(* IEC 61131-3 sources: plcassist-cli/packages/volt-lsp-iec/test-corpus/lenze-mid/Device/Plc Logic/Application/Library Manager/L_OEEA_Library, 3.26.4.21 (Lenze), 23 files *)

(* ---- GVL_AXISSIM.gvl ---- *)
VAR_GLOBAL
	FEEDERAXIS : AXIS_REF_SIM := STRUCT(eTraversingRange := 1, lrCycleLength := 1000.0, lrFeedConstant := 1000.0, dwGearNumerator := 100, dwGearDenominator := 1, eMctrlMode := 0, wNoOfHTLPeriods := 128);
END_VAR

(* ---- GVL_VALIDATIONTEST.gvl ---- *)
VAR_GLOBAL
	SCEXECUTETIMEARRAY : scExecuteTimeArray;
	SCMACHINEDATA_BASE : scMachineData_base;
	SCPERFORMANCE_BASE : scPerformance_base;
	ULISTART : ULINT;
	ULIEND : ULINT;
	XPRODUCTIONACTIVE : BOOL := TRUE;
	FBMACHINEPERFORMANCE_BASE : L_OEEA_MachinePerformance_Base;
	FBDOWNTIME_BASE : L_OEEA_Downtime_base;
	FBSHIFTOEEHISTORYALL : L_OEEA_ShiftOEEHistory;
	FBSHIFTOEEHISTORY_BASE : L_OEEA_ShiftOEEHistory_Base;
	FBSHIFTDOWNTIMEHISTORY_BASE : L_OEEA_ShiftDowntimeHistory_base;
	SCPDINTERNAL_BASE : scInternalVar;
	SCPDSHIFTDAYINDEX : scPDShiftData;
	SCPDINTERNALDOWNTIME_BASE : scInternalDownVar;
	SCDOWNTIME_BASE : scDowntime_base;
	SCSHIFTDOWNTIMEHISTORY_BASE : ARRAY [1..3] OF scDowntime_base;
	SCSHIFTHISTORYALL : ARRAY [1..3] OF scPerformance;
	SCPDSHIFTHISTORY_BASE : scVisuShiftHistory_base;
	SCPDPRODUCTIONDATA : scInternalProductionData;
	SCSHIFTVALUES : scCurrentShiftValues;
END_VAR

(* ---- LINE_OEE_GVL_VAR.gvl ---- *)
VAR_GLOBAL
	UINOOFMACHINES : UINT := 60;
	UINOOFHISTORICALWEEKS : UINT := 4;
END_VAR

(* ---- VERSIONCONSTANTS.gvl ---- *)
VAR_GLOBAL
	GC_BYAMOUNTOFGENERALDATA : BYTE := 50;
	GC_BYAMOUNTDOWNTIMEERRORS : BYTE := 10;
	GC_IFILTERSAMPLES : INT := 20;
END_VAR

(* ---- CALENDAR_WEEK.fun ---- *)
FUNCTION CALENDAR_WEEK : UINT
VAR_INPUT
	DTEXTDT : DATE_AND_TIME;
END_VAR
END_FUNCTION

(* ---- EXECUTIONTIME.fun ---- *)
FUNCTION EXECUTIONTIME : BOOL
VAR_INPUT
	SFBSTR : STRING;
	ULISTART : ULINT;
	ULIEND : ULINT;
END_VAR
VAR_IN_OUT
	AEXECUTION : scExecuteTime;
END_VAR
END_FUNCTION

(* ---- L_OEEA_CUSTOMIZABLE_COPYSTRUCT.fun ---- *)
FUNCTION L_OEEA_CUSTOMIZABLE_COPYSTRUCT : BOOL
VAR_INPUT
	PBYSOURCE : POINTER TO BYTE;
	PBYTARGET : POINTER TO BYTE;
	UISIZESOURCE : UINT;
	UISIZETARGET : UINT;
END_VAR
END_FUNCTION

(* ---- LRAXISPOSCOUNT.fun ---- *)
FUNCTION LRAXISPOSCOUNT : LREAL
VAR_INPUT
	LRAXISPOS : LREAL;
END_VAR
VAR_IN_OUT
	SCAXISPOSCOUNT : scAxisPosCount;
END_VAR
END_FUNCTION

(* ---- GLOBALTEXTLIST.fb ---- *)
FUNCTION_BLOCK GLOBALTEXTLIST
VAR
	M_TEXTLISTFILE : STRING(255);
	_STNAMESPACE : STRING;
END_VAR
END_FUNCTION_BLOCK

(* ---- IMAGEPOOL_AXIS_REF_SIM.fb ---- *)
FUNCTION_BLOCK IMAGEPOOL_AXIS_REF_SIM
VAR
	M_STNAMESPACE : STRING(80);
	M_STHELPVARID : STRING;
	M_STHELPVARPATH : STRING(255);
	M_STHELP : STRING;
	M_REGISTERIMAGES : BOOL := TRUE;
END_VAR
END_FUNCTION_BLOCK

METHOD FB_INIT : BOOL
VAR_INPUT
	BINITRETAINS : BOOL;
	BINCOPYCODE : BOOL;
END_VAR
END_METHOD

METHOD FB_REINIT : BOOL
END_METHOD

METHOD FB_EXIT : BOOL
VAR_INPUT
	BINCOPYCODE : BOOL;
END_VAR
END_METHOD

(* ---- L_MC1A_BASICACTUATINGSPEED.fb ---- *)
FUNCTION_BLOCK L_MC1A_BASICACTUATINGSPEED
VAR_INPUT
	XREGULATORON : BOOL;
	XRESETERROR : BOOL;
	XSETDRIVEQSP : BOOL;
	XENABLESETVEL : BOOL;
	XINVERTDIRECTION : BOOL;
	LRSETVEL : LREAL := 300.0;
	LRSETACC : LREAL := 100.0;
	LRSETDEC : LREAL := 100.0;
END_VAR
VAR_OUTPUT
	XERROR : BOOL;
	XBUSY : BOOL;
	EERRORID : L_IE1A_ErrorID;
	XCOMMUNICATIONOK : BOOL;
	XAXISREADY : BOOL;
	XAXISENABLED : BOOL;
	XDRIVEWARNING : BOOL;
	XDRIVEERROR : BOOL;
	DWDRIVEERRORID : DWORD;
	XDRIVEQSPACTIVE : BOOL;
	LRACTVEL : LREAL;
	XDIRECTIONPOSITIVE : BOOL;
	XDIRECTIONNEGATIVE : BOOL;
	WDIGITALINPUTS : WORD;
END_VAR
VAR_IN_OUT
	AXIS : AXIS_REF_SIM;
END_VAR
VAR
	L_TB1A_PT1FILTER1 : L_TB1A_PT1Filter := STRUCT(lrFilterTime := 0.02);
	L_MC1A_INTEGRATEAXIS1 : L_MC1A_IntegrateAxis;
	L_MC1A_DIFFERENTIATE2 : L_MC1A_Differentiate;
	L_MC1A_CONVX1 : L_MC1A_ConvX := STRUCT(diDenom := 1000000000);
	L_MC1A_CONVX2 : L_MC1A_ConvX;
	R_TRIG3 : R_TRIG;
	TON0 : TON := STRUCT(IN := TRUE, PT := TIME#1m0s0ms);
	TON1 : TON;
	TP1 : TP;
	X1STCYCLE : BOOL := TRUE;
	BYINITCOUNTER : BYTE;
	LRTASKCYCLETIME : LREAL;
	DITASKCYCLETIME : DINT;
	XINIT : BOOL := TRUE;
	LRACTVEL_INTERNAL : LREAL;
	LRREVPERSEC : LREAL;
	LITMP1 : LINT;
	LITMP2 : LINT;
	LITMP3 : LINT;
	LITMP6 : LINT;
	LITMP7 : LINT;
	RRANDOMNUMBER : REAL;
	RTMP : REAL;
	RHEATSINKTEMPINT : REAL;
	RHEATSINKFILTERTIME : REAL := 73.7;
	RIXTLOADINT : REAL;
	RIXTLOADFILTERTIME : REAL := 43.3;
	RIXT2LOADINT : REAL;
	RIXT2LOADFILTERTIME : REAL := 37.3;
	LROPERATIONTIME : LREAL;
	LROPERATIONTIMECU : LREAL;
	LRMODULOCYCLELENGTH_INTERNAL : LREAL;
	DIMODULOCYCLELENGTH_INTERNAL : DINT;
	LRPOSTOUNITFACTOR : LREAL;
	LRTMPEE : LREAL;
	DWMODULOCYCLERESIDUAL : DWORD;
	DIHALFMODULOCYCLELENGTH : DINT;
	DWRESIDUAL : DWORD;
	DIACTPOS : DINT;
	DIACTPOSOLD : DINT;
	XRESADDACTCYCLE : BOOL;
	XRESSUBACTCYCLE : BOOL;
	DWHTLCOUNTERVALUE_INTERNAL : DWORD;
	DIDELTAPOS : DINT;
	DIINPUTOLD : DINT;
	DITMPEE : DINT;
END_VAR
END_FUNCTION_BLOCK

METHOD METH_RAMPGENERATOR : LREAL
VAR_INPUT
	LRSETVEL : LREAL;
	LRSETACC : LREAL;
	LRSETDEC : LREAL;
	LRACTVEL : LREAL;
	XLOADSTARTVEL : BOOL;
	LRSTARTVEL : LREAL;
END_VAR
END_METHOD

METHOD ACT_SDOEMULATION
END_METHOD

METHOD METH_RANDOM : REAL
VAR_INPUT
	RRANDOMNUMBER : REAL;
END_VAR
END_METHOD

(* ---- L_MC1A_CONVX.fb ---- *)
FUNCTION_BLOCK L_MC1A_CONVX
VAR_INPUT
	DIIN : DINT;
	DINUM : DINT := 1;
	DIDENOM : DINT := 1;
END_VAR
VAR_OUTPUT
	DIOUT : DINT;
	XLIMIT : BOOL;
END_VAR
VAR
	LIOUT : LINT;
	LIREMAINDER : LINT;
	LITMP : LINT;
	LIDENOMINATOR : LINT;
END_VAR
END_FUNCTION_BLOCK

(* ---- L_MC1A_DIFFERENTIATE.fb ---- *)
FUNCTION_BLOCK L_MC1A_DIFFERENTIATE
VAR_INPUT
	LRPOSITIONIN : LREAL;
	ETRAVERSINGRANGE : WORD;
	LRCYCLELENGTH : LREAL := 360.0;
END_VAR
VAR_OUTPUT
	LRVELOCITYOUT : LREAL;
	XERROR : BOOL;
END_VAR
VAR
	TON0 : TON := STRUCT(IN := TRUE, PT := TIME#1m0s0ms);
	X1STCYCLE : BOOL := TRUE;
	BYINITCOUNTER : BYTE;
	LRTASKCYCLETIME : LREAL;
	LRCYCLELENGTHINTERNAL : LREAL;
	LRPOSITIONINLIMITED : LREAL;
	LRPOSITIONINLIMITEDOLD : LREAL;
END_VAR
END_FUNCTION_BLOCK

METHOD METH_SHORTESTWAY : LREAL
VAR_INPUT
	LRSETPOS : LREAL;
	LRACTPOS : LREAL;
	LRCYCLELENGTH : LREAL;
END_VAR
END_METHOD

(* ---- L_MC1A_INTEGRATEAXIS.fb ---- *)
FUNCTION_BLOCK L_MC1A_INTEGRATEAXIS
VAR_INPUT
	LRVELIN : LREAL;
	XLOADSTARTPOSITION : BOOL;
	LRSTARTPOSITION : LREAL;
	LRCYCLELENGTH : LREAL;
END_VAR
VAR_OUTPUT
	LRPOSOUT : LREAL;
	LRVELOUT : LREAL;
	XZEROCW : BOOL;
	XZEROCCW : BOOL;
	XZERO : BOOL;
END_VAR
VAR
	TON0 : TON := STRUCT(IN := TRUE, PT := TIME#1m0s0ms);
	X1STCYCLE : BOOL := TRUE;
	BYINITCOUNTER : BYTE;
	LRTASKCYCLETIME : LREAL;
	LRPOSOUT_OLD : LREAL;
END_VAR
END_FUNCTION_BLOCK

METHOD METH_ADDOFFSETCYCLIC : LREAL
VAR_INPUT
	LRSETPOS : LREAL;
	LRSETOFFSET : LREAL;
	LRCYCLELENGTH : LREAL;
END_VAR
END_METHOD

(* ---- L_OEEA_BASE_FBS.fb ---- *)
FUNCTION_BLOCK L_OEEA_BASE_FBS EXTENDS L_OEEA_FBs_COMMON
VAR_IN_OUT
	SCMACHINEDATA_BASE : scMachineData_base;
	SCPERFORMANCE_BASE : scPerformance_base;
	SCDOWNTIME_BASE : scDowntime_base;
END_VAR
VAR
	FBMACHINEPERFORMANCE : L_OEEA_MachinePerformance_Base;
	SCMACHINEDATA : scMachineData;
	FBDOWNTIME : L_OEEA_Downtime_Base;
	SCDOWNTIME : scDowntime;
END_VAR
END_FUNCTION_BLOCK

METHOD ACT_02_PRODUCTIONSIMULATIONSETTINGS
END_METHOD

METHOD ACT_12_CALL_MACHINEPERFORMANCE
END_METHOD

METHOD ACT_00_BASE_CONVERSION
END_METHOD

METHOD ACT_01_STANDARDASSIGNMENTS
END_METHOD

METHOD ACT_11_BREAKASSIGNMENTS
END_METHOD

METHOD ACT_10_SCHEDULERSELECTION
END_METHOD

(* ---- L_OEEA_FBS.fb ---- *)
FUNCTION_BLOCK L_OEEA_FBS EXTENDS L_OEEA_FBs_COMMON
VAR_IN_OUT
	SCMACHINEDATA : scMachineData;
	SCPERFORMANCE : scPerformance;
	SCACTUALSTATEDURATION : scVisuProductionStatus_base;
	SCDOWNTIME : scDowntime;
	SCVISU_IN_X_TREND : scXAxis_Trend;
	SCVISU_IN_Y_TREND : scYAxis_Trend;
	SCVISU_TREND_Y_LIMITS : scTrend_Limits;
END_VAR
VAR
	FBMACHINEPERFORMANCE : L_OEEA_MachinePerformance;
	FBDOWNTIME : L_OEEA_Downtime;
	FB_X_AXIS_TREND : L_OEEA_X_TREND;
	FB_Y_AXIS_TREND : L_OEEA_Y_TREND;
	XSORTUPDOWN : BOOL := TRUE;
	FBTIMETRIGGER : TON;
	FBTIMETRIGGER2 : TON;
	TXYGRAPHTIME : TIME := TIME#1m0s0ms;
	SPOWERUPJSONSUBSTR : STRING(255);
	ISETCALCTHROUGHPUT : INT;
	TSETTIMEXYGRAPH : TIME;
END_VAR
END_FUNCTION_BLOCK

METHOD ACT_01_STANDARDASSIGNMENTS
END_METHOD

METHOD ACT_13_CALL_PRODUCTION_TRENDS
END_METHOD

METHOD ACT_02_PRODUCTIONSIMULATIONSETTINGS
END_METHOD

METHOD ACT_12_CALL_MACHINEPERFORMANCE
END_METHOD

METHOD ACT_11_BREAKASSIGNMENTS
END_METHOD

METHOD ACT_10_SCHEDULERSELECTION
END_METHOD

(* ---- L_OEEA_FBS_COMMON.fb ---- *)
FUNCTION_BLOCK L_OEEA_FBS_COMMON
VAR_INPUT
	XENABLED : BOOL;
	XRESETACTUALDATA : BOOL;
	XRESETHISTORYDATA : BOOL;
	XPRODSIMULTIONENABLED : BOOL;
	XPRODSIMEVENTOCCURRENCE : BOOL := TRUE;
	XPRODSIMMATERIALPRODUCTION : BOOL;
	XHMIACTIVE : BOOL;
	ESCHEDULERMODE : L_OEEA_BaseDependency.enumShiftMode;
	ESETWEEKDAY : RTCLK.WEEKDAY;
	XDEACTIVESHIFTCONTINIOUSUPDATE : BOOL;
	UIMAXSIMULATIONEVENTS : UINT := 1;
	SCTRIGGER : scTrigger;
	XUSERESONCODESTRING : BOOL;
	XUPDATEJSONOEEKPI : BOOL;
	XMANUALSHIFTRESET : BOOL;
	XSHIFTPRODUCTIONACTIVE : BOOL;
	XLATERSHIFTSTARTENABLED : BOOL;
	SCSIMULATIONMODES : scSimulationModes;
	SREASONTEXTPOWERON : STRING := '';
END_VAR
VAR_OUTPUT
	XBUSY : BOOL;
	XERROR : BOOL;
	SCSHIFTVALUES : L_OEEA_ShiftScheduler.scCurrentShiftValues;
END_VAR
VAR_IN_OUT
	SCPRODUCTIONMODE : scProductionMode;
	ASERRORCATEGORY : scCategoryStruct;
	SCFIRSTERRORDATA : scErrorData;
	ASCDAYSCHEDULES : ARRAY [1..uiDaySchedule] OF scDaySchedule;
	SCPDINTERNAL : scInternalVar;
	SCPDINTERNALDOWNTIME : scInternalDownVar;
	SCPDPRODUCTIONDATA : scInternalProductionData;
	SCPDSHIFTDAYINDEX : scPDShiftData;
	SCPDSHIFTHISTORY_BASE : scVisuShiftHistory_base;
	SCSHIFTDOWNTIMEHISTORY : ARRAY [1..3] OF scDowntime_base;
	SCOEE_VISUPD : scOEE_VisuPD;
	SCVISU_OUT_PARTCORRECTION : scPartCorrectionInput;
	SCVISU_OUT_BUTTONS : scVisuButtons;
	SCSIMULATIONDOWNTIMES : scSimulationDowntimes;
END_VAR
VAR
	FBOEEA_SIMULATIONSETTINGS : L_OEEA_SimulationSettings;
	FBPRODUCTIONSCHEDULER : L_OEEA_ProductionScheduler;
	SCCUTREAL : scCutAverageReal;
	FBSHIFTCALENDAR : L_OEEA_ShiftScheduler.L_OEEA_ShiftScheduler;
	FBSTANDARDASSIGNMENT : L_OEEA_StandardAssignment;
	FBSHIFTOEEHISTORY : L_OEEA_ShiftOEEHistory_base;
	EPRODLOGFORMAT : eProduction_log := eProduction_log.Json;
	FBSHIFTDOWNTIMEHISTORY : L_OEEA_ShiftDowntimeHistory_base;
	XFIRSTCYCLE : BOOL := FALSE;
	XGETDEACTIVESHIFTCONTINIOUSUPDATE : BOOL;
	SSHIFTNAME : STRING;
	ICALCTHROUGHPUT : INT := 0;
	XRESETPRODLOGSHIFTCHANGE : BOOL;
	XFIRSTPLCCYCLEPROLONG : BOOL;
	SETSHIFTNAME : scShiftName;
END_VAR
END_FUNCTION_BLOCK

(* ---- L_OEEA_LINE_FB.fb ---- *)
FUNCTION_BLOCK L_OEEA_LINE_FB
VAR_INPUT
	XENABLE : BOOL;
	XRESETHISTORY : BOOL;
	UIMAXNOOFMACHINES : UINT;
	UINOOFCONNCTEDMACHINES : UINT;
	UINOOFHISTORICALWEEKS : UINT;
	TSETTIMEDEVIATION : TIME := TIME#10s0ms;
	TSETTIMECONNECTION : TIME := TIME#1m30s0ms;
	TSETTIMESHIFTCHANGEDELAY : TIME := TIME#5s0ms;
	TSETTIMELINEOEEUPDATEDELAY : TIME := TIME#10s0ms;
	SCTRIGGER : scTrigger_base;
	SCMACHINEOFFMODE : scMachineOffMode;
	SSHIFTNAME : STRING;
	ILINEID : INT;
	SLINEID : STRING;
END_VAR
VAR_OUTPUT
	XBUSY : BOOL;
	XDONE : BOOL;
	XERROR : BOOL;
	SCLINESTATUS : scLineStatus;
	XSHIFTCHANGEDELAYPROLONGTIME : BOOL;
	XLINEOEEUPDATEDELAYPROLONGTIME : BOOL;
	XLINEOEESTORAGEDELAY : BOOL;
END_VAR
VAR_IN_OUT
	ASCMACHINEDATA_NVL : ARRAY [1..Line_OEE_GVL_Var.uiNoOfMachines] OF scMachineData_NVL;
	ASCNVL : ARRAY [1..Line_OEE_GVL_Var.uiNoOfMachines] OF scRef_NVL;
	SCSHIFTVALUES : scCurrentShiftValues;
	SCLINEKPIS : scLineKPIs;
	ASCHISTORICALLINEKPIS : ARRAY [1..Line_OEE_GVL_Var.uiNoOfHistoricalWeeks] OF scLineKPIs;
	SCACTIVEDURINGACTUALSHIFT : ARRAY [1..Line_OEE_GVL_Var.uiNoOfMachines] OF scMachineShiftActive;
END_VAR
VAR
	I : INT;
	K : INT;
	N : INT;
	SCLINEKPISDEL : scLineKPIs;
	SCLINESTATUSDEL : scLineStatus;
	ROEE_WEIGHT : REAL;
	ROEERT : REAL;
	RTEEP : REAL;
	SLASTDATETIME : STRING;
	DTLASTDATETIME : DATE_AND_TIME;
	ISTRPOSBLANK : INT;
	TDATETIMEDIFF : TIME;
	XFIRSTNOTCONNECTEDMACHINE : BOOL;
	XFIRSTMACHINEDATETIMEINSYNCH : BOOL;
	XFIRSTNOTACTIVEMACHINE : BOOL;
	DTSHIFTSTART : DATE_AND_TIME;
	IWEEKDAYSDIFF : INT;
	DTDIFFSTARTTIME : TIME;
	DTPREVIOUSDATETIME : DATE_AND_TIME;
	TONPROLONGTIMER : ARRAY [1..2] OF TON;
	ISTEPSHIFTCHANGE : INT := 0;
	XSHIFTCHANGELINECONTROLLERDETECTED : BOOL;
	ILASTNOMACHINEACTIVEOEECALC : INT;
	SCDELACTIVEDURINGACTUALSHIFT : ARRAY [1..Line_OEE_GVL_Var.uiNoOfMachines] OF scMachineShiftActive;
END_VAR
END_FUNCTION_BLOCK

METHOD ACT_LINEOEEHISTORY
END_METHOD

METHOD ACT_CAL_OEEKPIS
END_METHOD

METHOD ACT_SHIFTSTARTTIME
END_METHOD

METHOD SUB_01_INIT_LOOP
END_METHOD

METHOD SUB_02_CHECK_STATUS
END_METHOD

METHOD SUB_03_CALC_MACHINEOEE
END_METHOD

METHOD SUB_04_CALC_LINEOEESUMMARY
END_METHOD

METHOD SUB_05_CALC_AVERAGELINEOEE
END_METHOD

METHOD SUB_06_SET_LINESTATUS
END_METHOD

METHOD METH_PROLONGBIT : BOOL
VAR_INPUT
	TPROLONGTIME : TIME;
END_VAR
VAR_IN_OUT
	TONPROLONGTIMER : TON;
	XSTARTPROLONGTIME : BOOL;
END_VAR
END_METHOD

METHOD ACT_SHIFTCHANGESEQ
END_METHOD

(* ---- L_OEEA_SIMULATIONAXIS.fb ---- *)
FUNCTION_BLOCK L_OEEA_SIMULATIONAXIS
VAR_INPUT
	XENABLED : BOOL;
	XDOWNTIMESTOP : BOOL;
	RTECHNICALCYCLETIME : REAL;
END_VAR
VAR_OUTPUT
	XMANUALSTOP : BOOL;
END_VAR
VAR_IN_OUT
	LRAXESACTMETERS : LREAL;
	LRAXESACTSCAPMETERS : LREAL;
END_VAR
VAR
	AXISJOG : L_MC1A_BasicActuatingSpeed;
	XREGULATORON : BOOL;
	XMOVEVELEXECUTE : BOOL;
	XJOGPOS : BOOL;
	XSTOP : BOOL;
	LRJOGGINGSETVEL : LREAL;
	ISTEP : INT;
	RFACTORPERFORMANCELOSS : REAL := 1.025;
	LRACTUALINCPOSITIONSIM : LREAL;
	LRACTUALDIFF : LREAL;
	TSCRAPMATERIALSTART : TON_Pausable;
	TSCRAPMATERIALSTOP : TON_Pausable;
END_VAR
END_FUNCTION_BLOCK

METHOD ACTMOTIONCTRL
END_METHOD

METHOD ACT_CALLMOTIONFB
END_METHOD

(* ---- L_OEEA_SIMULATIONSETTINGS.fb ---- *)
FUNCTION_BLOCK L_OEEA_SIMULATIONSETTINGS
VAR_INPUT
	XPRODSIMULTIONENABLED : BOOL;
	XPRODSIMEVENTOCCURRENCE : BOOL := TRUE;
	XRESETACTUALDATA : BOOL;
	ESCHEDULERMODE : enumShiftMode;
	XMATERIALPRODUCTION : BOOL;
	UIMAXSIMULATIONEVENTS : UINT := 1;
	SCSIMULATIONMODES : scSimulationModes;
END_VAR
VAR_OUTPUT
	XBUSY : BOOL;
	XERROR : BOOL;
END_VAR
VAR_IN_OUT
	SCMACHINEDATA : scMachineData;
	SCSHIFTVALUES : L_OEEA_ShiftScheduler.scCurrentShiftValues;
	SCDOWNTIME : scDowntime;
	SCSIMULATIONDOWNTIMES : scSimulationDowntimes;
	SCPRODUCTIONMODE : scProductionMode;
END_VAR
VAR
	SCRT_STATUS : RT_Status_Struct;
	FBDATASIMULATOR : L_OEEA_DataSimulator;
	XSTATIONENABLED : BOOL := TRUE;
	SCRT_STATUS_RESET : RT_Status_Struct;
	PA_TIMER : RT_Timer;
	PA_DOWNTIME : RT_Downtime;
	SCCUTREAL : scCutAverageReal;
	XFIRSTCYCLESIM : BOOL := FALSE;
	FBXHOLDINGACTIVE : R_TRIG;
	DILASTTYPEID : INT;
	IMAXSIMULATIONERRORS : INT;
	FBSIMULATIONAXIS : L_OEEA_SimulationAxis;
	XMANUALSTOP : BOOL;
	LRCOUNTOK : LREAL;
	LRCOUNTNOK : LREAL;
END_VAR
END_FUNCTION_BLOCK

METHOD ACT_03_MASCHINEPERFORMANCESIMULATION
END_METHOD

METHOD ACT_01_PRODUCTIONSIMULATION
END_METHOD

METHOD ACT_02_CALL_PRODUCTIONSIMULATOR
END_METHOD

METHOD ACT_04_CALLSIMULATIONAXIS
END_METHOD

(* ---- L_OEEA_STANDARDASSIGNMENT.fb ---- *)
FUNCTION_BLOCK L_OEEA_STANDARDASSIGNMENT
VAR_INPUT
	ENABLED : BOOL;
	XHMIACTIVE : BOOL;
END_VAR
VAR_OUTPUT
	XBUSY : BOOL;
	XERROR : BOOL;
END_VAR
VAR_IN_OUT
	SCSHIFTVALUES : L_OEEA_ShiftScheduler.scCurrentShiftValues;
	SCMACHINEDATA : scMachineData;
	SCDOWNTIME : scDowntime;
	SCPRODUCTIONMODE : scProductionMode;
	ASERRORCATEGORY : scCategoryStruct;
	SCFIRSTERRORDATA : scErrorData;
	ASCDAYSCHEDULES : ARRAY [1..uiDaySchedule] OF scDaySchedule;
	SCOEE_VISUPD : scOEE_VisuPD;
	SCVISU_OUT_BUTTONS : scVisuButtons;
	SCVISU_OUT_PARTCORRECTION : scPartCorrectionInput;
END_VAR
VAR
	I : INT;
	K : INT;
	IDEFAULTDAYOFWEEK : INT;
	IACTUALDAYOFWEEK : INT;
	XFIRSTCYCLE : BOOL := FALSE;
	FBXSAVESHIFTDATA : R_TRIG;
	ACTUALDAYINDEX : INT;
END_VAR
END_FUNCTION_BLOCK

METHOD ACT_01_PRODUCTIONMODES
END_METHOD

METHOD ACT_02_SETSHIFTINTERVALS
END_METHOD

METHOD ACT_03_MACHINEPERFORMANCESETTINGS
END_METHOD

(* ---- L_OEEA_VALIDATION_FBS.fb ---- *)
FUNCTION_BLOCK L_OEEA_VALIDATION_FBS EXTENDS L_OEEA_FBs
VAR
	FBPRODUCTIONSCHEDULER2 : L_OEEA_ProductionScheduler;
END_VAR
END_FUNCTION_BLOCK

METHOD ACT_12X_CALL_MACHINEPERFROMANCETEST
END_METHOD

(* ---- L_TB1A_PT1FILTER.fb ---- *)
FUNCTION_BLOCK L_TB1A_PT1FILTER
VAR_INPUT
	LRIN : LREAL;
	LRFILTERTIME : LREAL := 0.1;
END_VAR
VAR_OUTPUT
	LROUT : LREAL;
END_VAR
VAR
	TON0 : TON := STRUCT(IN := TRUE, PT := TIME#1m0s0ms);
	X1STCYCLE : BOOL := TRUE;
	BYINITCOUNTER : BYTE;
	LRTASKCYCLETIME : LREAL;
END_VAR
END_FUNCTION_BLOCK
